// TIA Portal V20 export
DATA_BLOCK "T3_Resultado"   // DB40940
{ S7_Optimized_Access := 'TRUE' }
AUTHOR : IA
FAMILY : PRUEBA
VERSION : 0.1
// Prueba IA 3: un Bool por prueba
// stored: AutoNumber false
   VAR
      OR_ok : Bool;   // T3_OR
      Ramas_ok : Bool;   // T3_Ramas
      Mul_ok : Bool;   // T3_Mul
      Div_ok : Bool;   // T3_Div
      Le_ok : Bool;   // T3_Le
      Ret_A_ok : Bool;   // T3_Ret_A
      Ret_B_ok : Bool;   // T3_Ret_B
      EqString_ok : Bool;   // T3_Eq_String
      Vida_OB126 : DInt;   // Sube 1 en cada ciclo si el OB126 se ejecuta
   END_VAR
BEGIN
END_DATA_BLOCK
